Fanuc KAREL source: KT00735.KL

PROGRAM KT00735
%NOLOCKGROUP
VAR
  ARG: ARRAY[4] OF BOOLEAN
  OUT: INTEGER
BEGIN
  OUT = ARRAY_LEN(ARG)
END KT00735
